# EPICS substitutions: iocs/motor/micos-ioc/db/MoCo.substitutions
# C's iocMicos MoCo.substitutions, P from st.cmd.
file "$(MOTOR)/db/motor.db"
{
pattern
{N, M,       DTYP,         C, S, DESC,         EGU,     DIR, VELO, VBAS, ACCL, BDST, BVEL, BACC, MRES, PREC, DHLM, DLLM, INIT}
{1, "m$(N)", "Micos MoCo", 0, 0, "motor $(N)", degrees, Pos, 1,    .1,   .2,   0,    1,    .2,   0.01, 5,    100,  -100, ""}
{2, "m$(N)", "Micos MoCo", 0, 1, "motor $(N)", degrees, Pos, 1,    .1,   .2,   0,    1,    .2,   0.01, 5,    100,  -100, ""}
}
